Staubli VAL3: dioItem.dtx

public string sComment
public dio dDio
